Fanuc KAREL source: KT00321.KL

PROGRAM KT00321
%NOLOCKGROUP
VAR
  P1: XYZWPREXT
  P2: XYZWPREXT
  OUT: BOOLEAN
BEGIN
  P1.X = 1.0
  P2.Y = 2.0
  P1.X = 1.0
  P2.Y = 2.0
  OUT = P1 <> P2
END KT00321
